PROGRAM MAIN
VAR
	PlcFirstCycle : BOOL := TRUE;
	
	Home : fbHome;

END_VAR
VAR CONSTANT
	ShutterCleanCmdEvent : stShutterCmdEvent := (
        Execute := FALSE,
        Cmd := ( CmdType := eShutterCmdType.NONE, Position := (Height := 0, Angle := 0 ) ) );
END_VAR


IF PlcFirstCycle THEN
	// Place for code done in first plc cycle
	
	PlcFirstCycle := FALSE;
END_IF

Home();

END_PROGRAM

(* stored: Version 1.1.0.1
   POU MAIN: Id {b477ade9-5e41-44da-827a-03687596879d}, SpecialFunc None *)
